(* IEC 61131-3 sources: nautilus/examples/remote-fleet/sites/well-2, 3 files *)

(* ---- types.st ---- *)
(* A root .st file with no PROGRAM is a project library, in scope for
   every task's compile — see docs/functions.md "A .ld library" (the same
   rule, one language over). Pump is the SAME shape scada/sites.yaml
   declares as its shared Template for all three sites, but this copy, not
   a shared package, is what ships: each site deploys alone. *)
TYPE
  Pump : STRUCT
    Run     : BOOL;   (* running feedback *)
    Fault   : BOOL;   (* VFD fault *)
    SpeedHz : LREAL;  (* actual speed *)
    SpeedSP : LREAL;  (* operator/SCADA setpoint — written locally or by
                         a Sparkplug NCMD member write from the SCADA host *)
  END_STRUCT;
END_TYPE

(* ---- sim.st ---- *)
(* Bench-only plant for well-2: a smaller wet well than well-1's (a
   different span calibration) and a smaller pump (a lower max flow). *)
PROGRAM Sim
VAR_EXTERNAL
    WellLevel      : LREAL;
    InflowLps      : LREAL;
    Pump1          : Pump;
    Pump1_RunCmd   : BOOL;
    Pump1_SpeedCmd : LREAL;
    SimDtS         : LREAL;
END_VAR
VAR
    outflowLps : LREAL;
    tSec       : LREAL;
END_VAR
VAR CONSTANT
    InflowVaryFrac : LREAL := 0.20;
    InflowPeriodS  : LREAL := 150.0;
    TwoPi          : LREAL := 6.2831853;
END_VAR

tSec := tSec + SimDtS;

IF Pump1_RunCmd THEN
    Pump1.SpeedHz := LIMIT(0.0, Pump1.SpeedHz + LIMIT(-10.0 * SimDtS, Pump1_SpeedCmd - Pump1.SpeedHz, 10.0 * SimDtS), 55.0);
ELSE
    Pump1.SpeedHz := MAX(0.0, Pump1.SpeedHz - 10.0 * SimDtS);
END_IF;
Pump1.Run := Pump1.SpeedHz > 5.0;
Pump1.Fault := FALSE;

(* ~0 below 30 Hz, 8 L/s at 55 Hz — a smaller pump than well-1's. *)
IF Pump1.SpeedHz <= 30.0 THEN
    outflowLps := 0.0;
ELSE
    outflowLps := (Pump1.SpeedHz - 30.0) / (55.0 - 30.0) * 8.0;
END_IF;

(* 1100 L span over 100 % (11 L per %) — a smaller wet well than well-1's. *)
WellLevel := LIMIT(0.0, WellLevel + (InflowLps * (1.0 + InflowVaryFrac * SIN(tSec / InflowPeriodS * TwoPi)) - outflowLps) * SimDtS / 11.0, 100.0);
END_PROGRAM

(* ---- well.st ---- *)
(* well-2's own control: the same shape as ../well-1/well.st, deliberately
   duplicated rather than shared — each site in this fleet deploys alone.
   Different setpoints live in this project's nautilus.yaml. *)
PROGRAM Well
VAR_EXTERNAL
    WellLevel     : LREAL;
    Pump1         : Pump;
    Pump1_RunCmd  : BOOL;
    Pump1_SpeedCmd : LREAL;
    PumpOnLevel   : LREAL;
    PumpOffLevel  : LREAL;
    MinSpeedHz    : LREAL;
    MaxSpeedHz    : LREAL;
    PumpStarts    : INT;
    PumpHours     : LREAL;
    WellDtS       : LREAL;
END_VAR
VAR
    edgeUp : R_TRIG;
END_VAR

Pump1_RunCmd := (WellLevel >= PumpOnLevel) OR (Pump1_RunCmd AND WellLevel > PumpOffLevel);

IF Pump1_RunCmd THEN
    Pump1_SpeedCmd := LIMIT(MinSpeedHz, Pump1.SpeedSP, MaxSpeedHz);
ELSE
    Pump1_SpeedCmd := 0.0;
END_IF;

edgeUp(CLK := Pump1.Run);
IF edgeUp.Q THEN
    PumpStarts := PumpStarts + 1;
END_IF;
IF Pump1.Run THEN
    PumpHours := PumpHours + WellDtS / 3600.0;
END_IF;
END_PROGRAM
